// TIA Portal V21 export
// export: Created 2026-08-21T20:18:54.7056607Z, ExportSetting None, DisplayName Totally Integrated Automation Portal, DisplayVersion V21, DisplayName STEP 7 Professional, DisplayVersion V21, DisplayName STEP 7 Safety, DisplayVersion V21, DisplayName Tech WebApplication, DisplayVersion V21, DisplayName WinCC Basic/Comfort/Advanced, DisplayVersion V21, DisplayName WinCC Professional, DisplayVersion V21, DisplayName WinCC Unified, DisplayVersion V21
TYPE "UDT_MTP_DIntProcessValueIn"
   STRUCT
      WQC { ExternalWritable := 'False'} : Byte := 16#FF;   // Worst Quality Code
      OSLevel : Byte;   // OSLevel variable
      V : DInt;   // Value
      VQC : Byte := 16#FF;   // Quality Code of the current received value
      SclMinCur { ExternalWritable := 'False'} : DInt;   // Value Scale Low Limit
      SclMaxCur { ExternalWritable := 'False'} : DInt := 100;   // Value Scale High Limit
      UnitCur { ExternalWritable := 'False'} : Int := 1998;   // Value Unit
      SclMinExt : DInt;   // External configuration for VScaleMin; If written value is valid VScaleMin will be set to VSclMinExt; If written value is invalid VScaleMin will be set to a predefined Value
      SclMaxExt : DInt := 100;   // External configuration for VScaleMax; If written value is valid VScaleMax will be set to VSclMaxExt; If written value is invalid VScaleMax will be set to a predefined Value
      UnitExt : Int := 1998;   // External configuration for VUnit; If written value is valid VUnit will be set to VUnitExt
      Apply : Bool;   // Apply new *Ext values to *Cur values
      ApplyEn { ExternalWritable := 'False'} : Bool;   // Flag to signalize if a new values can be applied; 1: new values can be applied; 0: currently, no new value can be applied
   END_STRUCT;
END_TYPE
